// TIA Portal V21 export
// export: Created 2026-11-07T15:50:59.4306851Z, ExportSetting WithDefaults, DisplayName Totally Integrated Automation Portal, DisplayVersion V21, DisplayName STEP 7 Professional, DisplayVersion V21, DisplayName STEP 7 Safety, DisplayVersion V21, DisplayName Tech WebApplication, DisplayVersion V21, DisplayName WinCC Basic/Comfort/Advanced, DisplayVersion V21, DisplayName WinCC Unified, DisplayVersion V21
TextList "TL_Alarm"  ListRange=Decimal
  TextListEntry   EntryType=SingleValue, From=-1, To=-1, Text="-"
  TextListEntry   EntryType=SingleValue, Text="0 Neuravnoteženost broda |L-R| > 5"
  TextListEntry   EntryType=SingleValue, From=1, To=1, Text="1 Lokacija podizanja prazna"
  TextListEntry   EntryType=SingleValue, From=2, To=2, Text="2 Lokacija spuštanja zauzeta"
  TextListEntry   EntryType=SingleValue, From=3, To=3, Text="3 ID u listi za istovar, nije u Bay 0"
  TextListEntry   EntryType=SingleValue, From=4, To=4, Text="4 ID u listi za ukrcaj, nije u Bay 1"
  TextListEntry   EntryType=SingleValue, From=5, To=5, Text="5 Neispravan ID (100-999)"
  TextListEntry   EntryType=SingleValue, From=6, To=6, Text="6 Dvostruki ID"
  TextListEntry   EntryType=SingleValue, From=7, To=7, Text="7 Nema slobodnog mjesta"
  TextListEntry   EntryType=SingleValue, From=8, To=8, Text="8 Plan nije izvediv"
  TextListEntry   EntryType=SingleValue, From=9, To=9, Text="9 Neispravna ručna naredba"
  TextListEntry   EntryType=SingleValue, From=10, To=10, Text="10 Dizalica: timeout naredbe"
  TextListEntry   EntryType=SingleValue, From=11, To=11, Text="11 Dizalica već nosi kontejner"
  TextListEntry   EntryType=SingleValue, From=12, To=12, Text="12 Dizalica ne nosi kontejner"
  TextListEntry   EntryType=SingleValue, From=13, To=13, Text="13 Nije inicijalizirano"
  TextListEntry   EntryType=SingleValue, From=14, To=14, Text="14 Položaj dizalice ne odgovara"
  TextListEntry   EntryType=SingleValue, From=15, To=15, Text="15 Istovar i ukrcaj završeni"
